(* IEC 61131-3 sources: kns-port-domestic/tools/plcopen/tests/fixtures/constructs/src/Interfaces/I_Resettable, 1 file *)

(* ---- Reset.method.decl.st ---- *)
// Сбросить; TRUE — сброс выполнен
METHOD Reset : BOOL
VAR_INPUT
    xForce : BOOL;
END_VAR
